(* PLC project , Example Fixture *)

PROGRAM Main
  VAR_INPUT
    Skip : BOOL;
    Start : BOOL;
  END_VAR
  VAR_OUTPUT
    Lamp : BOOL;
  END_VAR

(* LD diagram, written out as Structured Text *)
IF Skip THEN JMP Over; END_IF;
Lamp := Start;
Over:
END_PROGRAM

CONFIGURATION c
  RESOURCE r ON PLC
    TASK t(INTERVAL := T#10ms, PRIORITY := 1);
    PROGRAM t_i WITH t : Main;
  END_RESOURCE
END_CONFIGURATION
